// TIA Portal V21 export
// export: Created 2026-11-11T00:47:38.7533279Z, ExportSetting WithDefaults, DisplayName Totally Integrated Automation Portal, DisplayVersion V21 Update 3, DisplayName STEP 7 Professional, DisplayVersion V21 Update 3, DisplayName STEP 7 Safety, DisplayVersion V21, DisplayName Tech WebApplication, DisplayVersion V21, DisplayName WinCC Basic/Comfort/Advanced, DisplayVersion V21 Update 3, DisplayName WinCC Unified, DisplayVersion V21 Update 3
FUNCTION_BLOCK "FB_Fbd_ex147"   // FB155, FBD
{ S7_Optimized_Access := 'TRUE' }
VERSION : 0.1
// stored: AutoNumber true, IsIECCheckEnabled false, IsRetainMemResEnabled false, MemoryReserve 100, SetENOAutomatically false, UDAEnableTagReadback false
   VAR_INPUT
      v_req : Bool;
      v_low_limit : UInt;
      v_up_limit : UInt;
      v_count : UDInt;
      v_attrib : Byte;
      v_srcblk : Variant;
   END_VAR
   VAR_OUTPUT
      v_ret_val : Int;
      v_busy : Bool;
      v_db_num : UInt;
   END_VAR
BEGIN

REGION Network 1: CREATE_DB - Create data block
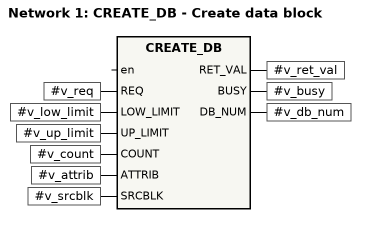
   #v_ret_val := CREATE_DB(REQ := #v_req,
                           LOW_LIMIT := #v_low_limit,
                           UP_LIMIT := #v_up_limit,
                           COUNT := #v_count,
                           ATTRIB := #v_attrib,
                           SRCBLK := #v_srcblk,
                           BUSY => #v_busy,
                           DB_NUM => #v_db_num);
END_REGION
END_FUNCTION_BLOCK
